Fanuc KAREL source: KB00125.KL

PROGRAM KB00125
%NOLOCKGROUP
%ENVIRONMENT FLBT
VAR
  P1: STRING[80]
  P2: INTEGER
BEGIN
  P1 = 'A'
  P2 = 1
  MSG_DISCO(P1, P2)
END KB00125
